{attribute 'qualified_only'}
VAR_GLOBAL
	
	fbIoOutGroup		: FB_IoGroup;


	
	{attribute 'TcLinkTo' := '._bHw  := TIID^Device 1 (EtherCAT)^Term 18 (EK1200)^Term 22 (EL2008)^Channel 1^Output'}
	Ledred1 : FB_IoOutput(fbIoOutGroup);
	
	{attribute 'TcLinkTo' := '._bHw  := TIID^Device 1 (EtherCAT)^Term 18 (EK1200)^Term 22 (EL2008)^Channel 2^Output'}
	Ledgreen1 : FB_IoOutput(fbIoOutGroup);
	
	{attribute 'TcLinkTo' := '._bHw  := TIID^Device 1 (EtherCAT)^Term 18 (EK1200)^Term 22 (EL2008)^Channel 3^Output'}
	Ledgreen2 : FB_IoOutput(fbIoOutGroup);
	
	{attribute 'TcLinkTo' := '._bHw  := TIID^Device 1 (EtherCAT)^Term 18 (EK1200)^Term 22 (EL2008)^Channel 4^Output'}
	Ledred2 : FB_IoOutput(fbIoOutGroup);
	
	{attribute 'TcLinkTo' := '._bHw  := TIID^Device 1 (EtherCAT)^Term 18 (EK1200)^Term 22 (EL2008)^Channel 5^Output'}
	Ledred3 : FB_IoOutput(fbIoOutGroup);
END_VAR

(* stored: Version 1.1.0.1
   GVL Out: Id {f5dcc463-15a3-4edc-9337-062b34989f62} *)
